Fanuc KAREL source: kt00535.KL

PROGRAM KT00535
%STACKSIZE=65535
%PRIORITY=65535
%NOLOCKGROUP
VAR
P1 : JOINTPOS9
P2 : POSITION
OUT : XYZWPR
BEGIN
-- UNRESOLVED_PC line 8 opcodes [49 7E 49 60 7E 4A] marker_code=0
END KT00535
